// TIA Portal V21 export
// export: Created 2026-11-08T21:17:26.2737961Z, ExportSetting WithDefaults, DisplayName Totally Integrated Automation Portal, DisplayVersion V21 Update 3, DisplayName STEP 7 Professional, DisplayVersion V21 Update 3, DisplayName STEP 7 Safety, DisplayVersion V21, DisplayName Tech WebApplication, DisplayVersion V21, DisplayName WinCC Basic/Comfort/Advanced, DisplayVersion V21 Update 3, DisplayName WinCC Unified, DisplayVersion V21 Update 3
DATA_BLOCK "DB_AllTypes"   // DB6
{ S7_Optimized_Access := 'TRUE' }
VERSION : 0.1
// stored: AutoNumber true, DBAccessibleFromOPCUA true, DBAccessibleFromWebserver true, IsOnlyStoredInLoadMemory false, IsRetainMemResEnabled false, IsWriteProtectedInAS false, MemoryReserve 100
   VAR
      vBool : Bool := TRUE;   // Bool comment
      vByte : Byte := 16#12;
   END_VAR
   VAR RETAIN
      vWord : Word := 16#1234;
   END_VAR
   VAR
      vDWord : DWord := 16#12345678;
      vLWord : LWord := 16#123456789ABCDEF0;
      vSInt : SInt := -12;
      vUSInt : USInt := 200;
      vInt { ExternalAccessible := 'False'; ExternalVisible := 'False'; ExternalWritable := 'False'} : Int := -1234;
      vUInt : UInt := 60000;
      vDInt { ExternalWritable := 'False'} : DInt := -123456;
      vUDInt : UDInt := 4000000000;
      vLInt : LInt := -9000000000;
      vULInt : ULInt := 18000000000;
      vReal { ExternalVisible := 'False'} : Real := 1.5;
      vLReal : LReal := -2.25;
      vS5Time : S5Time := S5T#2S;
      vTime : Time := T#1H2M3S;
      vLTime : LTime := LT#5MS;
      vDate : Date := D#2026-11-05;
      vTod : Time_Of_Day := TOD#12:34:56;
      vLTod : LTime_Of_Day := LTOD#01:02:03.5;
      vDt : Date_And_Time := DT#2026-11-05-12:00:00;
      vLdt : LDT := LDT#2026-11-05-12:00:00;
      vDtl : DTL;
      vChar : Char := 'A';
      vWChar : WChar := WCHAR#'Z';
      vString : String := 'hello';
      vString10 : String[10] := 'ten';
      vWString : WString := WSTRING#'wide';
      vWString5 : WString[5];
      vSetpoint : Int;
      aNeg : Array[-2..2] of Int;
      a2d : Array[0..2, 1..3] of Real;
      a3d : Array[0..1, 0..1, 0..1] of Bool;
      aStr : Array[0..1] of String[8];
      aStruct : Array[0..1] of Struct
         x : Int;
         y : Bool;
      END_STRUCT;
      aUdt { S7_SetPoint := 'True'} : Array[0..2] of "UDT_Inner";
      a2dUdt { S7_SetPoint := 'True'} : Array[0..1, 0..1] of "UDT_Outer";
      outer { S7_SetPoint := 'True'} : "UDT_Outer";
      deep : Struct
         l1 : Struct
            l2 : Struct
               v : LReal := 3.14;
               arr : Array[0..1] of Struct
                  z : Word;
               END_STRUCT;
            END_STRUCT;
         END_STRUCT;
      END_STRUCT;
      vTimer { S7_SetPoint := 'True'} : IEC_TIMER;
      vCounter { S7_SetPoint := 'True'} : IEC_COUNTER;
   END_VAR
   VAR RETAIN
      rCount : UDInt;   // Retain counter
      rArr : Array[0..3] of Real;
   END_VAR
BEGIN
   aNeg[2] := 20;
   aNeg[-2] := -20;
   a2d[1,2] := 1.25;
   a3d[1,1,1] := TRUE;
   aStr[1] := 'abc';
   aStruct[1].x := 7;
   aUdt[2].Temp := 99.5;
   a2dUdt[1,0].inner.Static := 5;
   outer.txt := 'changed';
   deep.l1.l2.arr[1].z := 16#BEEF;
   rArr[3] := 0.5;
END_DATA_BLOCK
